Staubli VAL3: HMI_cycle.pjx

--- HMI_cycle.pjx ---
Parameters version=s8.15.3Cs9_BS3337 stackSize=5000 millimeterUnit=true
Program file=_clickAlarmAck.pgx
Program file=bind.pgx
Program file=click_End.pgx
Program file=click_Hold.pgx
Program file=click_Reset.pgx
Program file=click_RotHome.pgx
Program file=click_Start.pgx
Program file=click_Stop.pgx
Program file=currentState.pgx
Program file=cycletime.pgx
Program file=main.pgx
Program file=start.pgx
Program file=stop.pgx
Data file=HMI_cycle.dtx
Library alias=util path=Disk://HMI_cs9/HMI_util/HMI_util.pjx
Library alias=rs path=Disk://source/projectSource/robotStatus/robotStatus.pjx
Library alias=simulate path=Disk://HMI_cs9/simulate/simulate.pjx
Library alias=saveData path=Disk://source/saveData/saveData.pjx

--- HMI_cycle.dtx ---
mdesc mNomSpeed
bool bReset
bool bStart
bool bHold
bool bEnd
bool bStop
bool bBack
bool bToHome
bool bClearErr
string sState
string sCapacity
string sAvgCapacity
string sBestCapacity
string sProgCode
num nLastProg
string sTrajStatus
string sLib
num nLastLib
bool bRotBack

--- main.pgx ---
public program main()
  local bool l_bExit
  local string l_sTColor
  local string l_sEColor
  local num l_nClock
  local string l_sFColor
begin
  do
    if util:sPage!="cycle"
      util:sPage="cycle"
      call util:loadingPage()
      call bind()
      userPage(util:sPage)
      delay(0.5)
      l_sTColor="#33FF33"
      l_sFColor="#FFFFFF"
      l_sEColor="#FF3366"
      nLastProg=-1
    endIf

    //机器人状态
    call currentState()
    //button
    if bReset
      bReset=false
      call click_Reset()
    elseIf bStart
      bStart=false
      call click_Start()
    elseIf bHold
      bHold=false
      call click_Hold()
    elseIf bEnd
      bEnd=false
      call click_End()
    elseIf bStop
      bStop=false
      call  click_Stop()
    elseIf bBack
      bBack=false
      l_bExit=true
    elseIf bToHome
      bToHome=false
      call simulate:simulateHome()
    elseIf bRotBack
      bRotBack=false
      call click_RotHome()
    elseIf bClearErr
      bClearErr=false
      call _clickAlarmAck()
    endIf
    //数据库显示
    //if saveData:nLibIndex!=nLastLib
    //nLastLib=saveData:nLibIndex
    sLib=toString("",saveData:nLibIndex)
    //endIf
    //程序号显示
    if rs:nProgCode!=nLastProg
      nLastProg=rs:nProgCode
      sProgCode=toString("",rs:nProgCode)
    endIf
    //cycletime
    call cycletime()
    //500ms refresh
    if clock()-l_nClock>0.5
      l_nClock=clock()
      sTrajStatus=rs:sTrajStatus
      if rs:bIsHome
        userPageSet("cycle","btn1","style.backgroundColor",l_sTColor)
      else
        userPageSet("cycle","btn1","style.backgroundColor",l_sFColor)
      endIf
      if rs:bIsEstop
        userPageSet("cycle","btn2","style.backgroundColor",l_sEColor)
      else
        userPageSet("cycle","btn2","style.backgroundColor",l_sFColor)
      endIf
      if rs:bIsCycle
        userPageSet("cycle","btn3","style.backgroundColor",l_sTColor)
      else
        userPageSet("cycle","btn3","style.backgroundColor",l_sFColor)
      endIf
      if rs:bIsReady
        userPageSet("cycle","btn4","style.backgroundColor",l_sTColor)
      else
        userPageSet("cycle","btn4","style.backgroundColor",l_sFColor)
      endIf
      if rs:_bHeavyAlarm
        userPageSet("cycle","btn4_Copy1","style.backgroundColor",l_sTColor)
      else
        userPageSet("cycle","btn4_Copy1","style.backgroundColor",l_sFColor)
      endIf
    endIf
    delay(0)
  until l_bExit==true
end

--- start.pgx ---
program start()
begin
end

--- _clickAlarmAck.pgx ---
program _clickAlarmAck()
begin
  rs:_sRobotStatus="收到页面点击清除报错!"
  rs:bAlarmAck=true
  delay(0.1)
  rs:bAlarmAck=false
end

--- bind.pgx ---
program bind()
begin
  userPageBindClick("cycle","btn5",bReset,true)
  userPageBindClick("cycle","btn6",bStart,true)
  userPageBindClick("cycle","btn7",bHold,true)
  userPageBindClick("cycle","btn8",bEnd,true)
  userPageBindClick("cycle","btn9",bStop,true)
  userPageBindClick("cycle","btn10",bToHome,true)
  userPageBindClick("cycle","btnback",bBack,true)
  userPageBindClick("cycle","btn6_Copy1",bClearErr,true)
  userPageBindClick("cycle","btnRotback",bRotBack,true)
  userPageBind("cycle","lblStatus","innerHTML",sTrajStatus,1,"r")
  userPageBind("cycle","lbl8","innerHTML",sCapacity,1,"r")
  userPageBind("cycle","lbl9","innerHTML",sAvgCapacity,1,"r")
  userPageBind("cycle","lbl10","innerHTML",sBestCapacity,1,"r")
  userPageBind("cycle","lbl10_Copy1","innerHTML",sLib,1,"r")
  userPageBind("cycle","lbl10_Copy3","innerHTML",sProgCode,1,"r")
  userPageBind("cycle","lbl3","innerHTML",sState,1,"r")


  userPageBind("cycle","lst1","options",rs:sAlarmMes,size(rs:sAlarmMes),"r")


end

--- click_End.pgx ---
program click_End()
  local bool l_bResult
begin
   //循环停止机器人
  l_bResult=userPageConfirm("确认循环停止机器人？")
  if l_bResult
    rs:nCycleCmd=5
    delay(0.2)
    rs:nCycleCmd=0
  endIf
end

--- click_Hold.pgx ---
program click_Hold()
  local bool l_bResult
begin
   //暂停机器人
  l_bResult=userPageConfirm("确认暂停机器人？")
  if l_bResult
    rs:bToPause=true
    delay(0.2)
    rs:bToPause=false
  endIf
end

--- click_Reset.pgx ---
program click_Reset()
  local bool l_bResult
begin
  //   //复位机器人
  //  l_bResult=userPageConfirm("确认复位机器人？")
  //  if l_bResult
  //    rs:nCycleCmd=1
  //    delay(0.2)
  //    rs:nCycleCmd=0
  //  endIf
end

--- click_RotHome.pgx ---
program click_RotHome()
  local bool l_bResult
begin
  if workingMode()!=1
    popUpMsg("非手动模式不支持路径回原！")
    return
  endIf
  //手动机器人路径回原
  l_bResult=userPageConfirm("确认原路径返回Home？")
  if l_bResult
    rs:nCycleCmd=7
    delay(0.2)
    rs:nCycleCmd=0
  endIf

end

--- click_Start.pgx ---
program click_Start()
  local bool l_bResult
begin
  //启动机器人
  l_bResult=userPageConfirm("确认启动机器人？")
  if l_bResult
    rs:bToStartCycle=true
    delay(0.2)
    rs:bToStartCycle=false
  endIf
end

--- click_Stop.pgx ---
program click_Stop()
  local bool l_bResult
begin
  //立即停止机器人
  l_bResult=userPageConfirm("确认立即停止机器人？")
  if l_bResult
    rs:bToStopCycle=true
    delay(0.2)
    rs:bToStopCycle=false
  endIf
end

--- currentState.pgx ---
program currentState()
begin
  switch rs:_nOmacStat
    case 1
      sState="准备就绪"
    break
    case 2
      sState="正在启动"
    break
    case 3
      sState="运行中"
    break
    case 4
      sState="复位中"
    break
    case 5
      sState="暂停中"
    break
     case 6
      sState="已暂停"
    break
    case 7
      sState="正在结束周期"
    break
    case 8
      sState="停止中"
    break
    case 9
      sState="已停止"
    break
    case 10
      sState="任务终止中"
    break

  endSwitch
end

--- cycletime.pgx ---
program cycletime()
  local num l_nTotleCT
  local num l_nElement
  local num l_n
begin
  if rs:_nOmacStat==3
    //cunrrent capacity
    if rs:_nCycleTime[rs:_nCTIndex]>0
      rs:_nCapacity=60/rs:_nCycleTime[rs:_nCTIndex]
    else
      rs:_nCapacity=0
    endIf
    //average capacity
    l_nTotleCT=0
    l_nElement=0
    for l_n=0 to size(rs:_nCycleTime)-1
      if rs:_nCycleTime[l_n]!=0
        l_nTotleCT=l_nTotleCT+rs:_nCycleTime[l_n]
        l_nElement=l_nElement+1
      endIf
    endFor
    if l_nTotleCT>0
      rs:_nAvgCapacity=60*l_nElement/l_nTotleCT
    else
      rs:_nAvgCapacity=0
    endIf
    //best capacity
    rs:_nBestCapacity=max(rs:_nBestCapacity,rs:_nCapacity)
  else
    rs:_nCapacity=0
    rs:_nAvgCapacity=0
    rs:_nBestCapacity=0
  endIf
  sCapacity=toString(".2",rs:_nCapacity)
  sAvgCapacity=toString(".2",rs:_nAvgCapacity)
  sBestCapacity=toString(".2",rs:_nBestCapacity)
end

--- stop.pgx ---
program stop()
begin
end
